(* IEC 61131-3 sources: JingjiangArm/moonboxpro_arm_8.4/Application/Application/任务列表/CommTask/COMM_DIAMONDS/和金刚UDP通讯/ModBus协议相关, 8 files *)

(* ---- StADU.st ---- *)
(*@CES
Name=StADU
Type=Gvl
TypeGuid=2db5746d-d284-4425-9f7f-2663a34b0ebc
Guid=730e2a17-289c-4459-a153-1a559c1b0add
HasDeclaration=True
HasImplementation=False
*)
{DECLARATION}
{attribute 'pack_mode' := '1'}
TYPE StADU :(*Modbus-UDP应用层协议的7个字节*)
STRUCT
	stStMBAP: StMBAP;(*ModBus Application Protocol*)
	stStPDU_Header: StPDU_Header;(*PDU基础头/主要针对03和16两个功能字的请求*)
END_STRUCT
END_TYPE

{IMPLEMENTATION}

(* ---- StDataNode.st ---- *)
(*@CES
Name=StDataNode
Type=Gvl
TypeGuid=2db5746d-d284-4425-9f7f-2663a34b0ebc
Guid=d2752c56-02c4-4ac3-a8e3-7575782c62c6
HasDeclaration=True
HasImplementation=False
*)
{DECLARATION}
{attribute 'pack_mode' := '1'}
TYPE StDataNode :(*Modbus读写区域*)
STRUCT
	uiAddress: UINT;(*寄存器地址/相对于字节数有2倍关系*)
	uiQuantity: UINT;(*寄存器数量*)
	bySynchronized: BYTE;(*同步过的标志/0表示未同步/1表示当前在fifo中/255表示已经完成同步*)
	xRd_ing: BOOL;(*写操作进行中*)
	xWr_ing: BOOL;(*读操作进行中*)
END_STRUCT
END_TYPE

{IMPLEMENTATION}

(* ---- StDataZone.st ---- *)
(*@CES
Name=StDataZone
Type=Gvl
TypeGuid=2db5746d-d284-4425-9f7f-2663a34b0ebc
Guid=9a2c4743-5919-4081-a37c-2820a2d84e25
HasDeclaration=True
HasImplementation=False
*)
{DECLARATION}
{attribute 'pack_mode' := '1'}
TYPE StDataZone :(*Modbus读写区域*)
(*读写区域/节点地址+PARAM_ZONE_ALTERNATE_OFST*)
(*只写区域/节点地址+PARAM_ZONE_C2S*)
STRUCT
	uiNodeNum: UINT;(*节点数量/最大65535*)
	astStDataNode: ARRAY [1..MAX_DATA_NODE_NUM] OF StDataNode;
END_STRUCT
END_TYPE

{IMPLEMENTATION}

(* ---- StMBAP.st ---- *)
(*@CES
Name=StMBAP
Type=Gvl
TypeGuid=2db5746d-d284-4425-9f7f-2663a34b0ebc
Guid=18e79d68-9469-4b38-b2f6-5459a353a7ac
HasDeclaration=True
HasImplementation=False
*)
{DECLARATION}
{attribute 'pack_mode' := '1'}
TYPE StMBAP :(*Modbus-UDP应用层协议的7个字节*)
STRUCT
	uiInvocation: UINT;(*调用操作标识*)
	uiProtocol: UINT;(*协议*)
	uiLength: UINT;(*数据长度*)
	byUnit: BYTE;(*远程单元标识*)
END_STRUCT
END_TYPE

{IMPLEMENTATION}

(* ---- StPDU_Header.st ---- *)
(*@CES
Name=StPDU_Header
Type=Gvl
TypeGuid=2db5746d-d284-4425-9f7f-2663a34b0ebc
Guid=e7e8d47d-075f-4d58-8263-79c4bddf08e0
HasDeclaration=True
HasImplementation=False
*)
{DECLARATION}
{attribute 'pack_mode' := '1'}
TYPE StPDU_Header :(*Modbus/功能码/起始地址/寄存器数量*)
STRUCT
	byFunction: BYTE;
	uiAddress: UINT;
	uiQuantity: UINT;
END_STRUCT
END_TYPE

{IMPLEMENTATION}

(* ---- StProofItem.st ---- *)
(*@CES
Name=StProofItem
Type=Gvl
TypeGuid=2db5746d-d284-4425-9f7f-2663a34b0ebc
Guid=570fb4d9-10a9-4892-8e2d-1d8339482480
HasDeclaration=True
HasImplementation=False
*)
{DECLARATION}
{attribute 'pack_mode' := '1'}
TYPE StProofItem :(*证据链*)
STRUCT
	iWaitRespCycles: INT;(*等待响应的周期次数/超时就把这个后面的报文重置/把该计数清零*)
	stStADU: StADU;(*发送的16功能字报文*)
END_STRUCT
END_TYPE

{IMPLEMENTATION}

(* ---- StProofList.st ---- *)
(*@CES
Name=StProofList
Type=Gvl
TypeGuid=2db5746d-d284-4425-9f7f-2663a34b0ebc
Guid=df0f82a0-67c4-4a3b-a0bd-b03f60b31cfe
HasDeclaration=True
HasImplementation=False
*)
{DECLARATION}
{attribute 'pack_mode' := '1'}
TYPE StProofList :(*证据链*)
STRUCT
	astStProofItem: ARRAY [1..MAX_MB_FIFO_ITEMS] OF StProofItem;
END_STRUCT
END_TYPE

{IMPLEMENTATION}

(* ---- StZone_W.st ---- *)
(*@CES
Name=StZone_W
Type=Gvl
TypeGuid=2db5746d-d284-4425-9f7f-2663a34b0ebc
Guid=aa2f6bf5-5ddf-4cba-b55b-f3a209fac971
HasDeclaration=True
HasImplementation=False
*)
{DECLARATION}
{attribute 'pack_mode' := '1'}
TYPE StZone_W :(*Modbus只写区域*)
(*节点地址+PARAM_ZONE_C2S*)
STRUCT
	stStMBAP: StMBAP;(*ModBus Application Protocol*)
	stStPDU_Header: StPDU_Header;(*PDU基础头/主要针对03和16两个功能字的请求*)
END_STRUCT
END_TYPE

{IMPLEMENTATION}
